TYPE ST_CameraProcessSettings :
STRUCT
    udiMovingTriggerDelayMs : UDINT := 100;
    udiRotaryConfirmMs : UDINT := 1000;
END_STRUCT
END_TYPE

(* stored: Version 1.1.0.1, ProductVersion 3.1.4026.18
   DUT ST_CameraProcessSettings: Id {a56202e9-5472-4e0b-84b7-8b2daa8ffbbd} *)
